(* IEC 61131-3 sources: PortalRobot/Portal_robot/Device/application/ST/ST_STATISTIC, 4 files *)

(* ---- ST_STATISTIC.st ---- *)
TYPE ST_STATISTIC :
STRUCT
	stMachineStat 		: ST_STATISTIC_MACHINE;
	stRobotStat 		: ST_STATISTIC_ROBOT;
END_STRUCT
END_TYPE

(* ---- ST_STATISTIC_MACHINE.st ---- *)
TYPE ST_STATISTIC_MACHINE :
STRUCT
	rLoadCNC_1            : REAL; // Процент загрузки станка 1
	rLoadCNC_2            : REAL; // Процент загрузки станка 2
	rLoadCNC_3            : REAL; // Процент загрузки станка 3
END_STRUCT
END_TYPE

(* ---- ST_STATISTIC_ROBOT.st ---- *)
TYPE ST_STATISTIC_ROBOT :
STRUCT
	tCNC_1      	: TIME; // Среднее время работы в стнке 1
	tCNC_2      	: TIME; // Среднее время работы в стнке 2
	tCNC_3      	: TIME; // Среднее время работы в стнке 3
	tMoveCNC_1 		: TIME; // Среднее время перемещения от магазина к станку 1
	tMoveCNC_2 		: TIME; // Среднее время перемещения от магазина к станку 2
	tMoveCNC_3 		: TIME; // Среднее время перемещения от магазина к станку 3
	tMagazine       : TIME; // Среднее время работы в магазине

	rRobot          : REAL; // Процент загрузки робота
END_STRUCT
END_TYPE

(* ---- ST_STATISTIC_SAMPLE.st ---- *)
TYPE ST_STATISTIC_SAMPLE :
STRUCT
    uliElapsedMs : ULINT; // Накопленное время сессии с учётом ускорения
    auliBusyMs : ARRAY [1..11] OF ULINT; // Завершённые и текущие интервалы
    auliCompletedBusyMs : ARRAY [1..11] OF ULINT; // Только завершённые интервалы
    auliCompletedCount : ARRAY [1..11] OF ULINT;
END_STRUCT
END_TYPE
